Fanuc KAREL source: KT00971.KL

PROGRAM KT00971
%NOLOCKGROUP
VAR
  ENTRY: INTEGER
  PNAME: STRING[80]
  VNAME: STRING[80]
  STATUS: INTEGER
  VALUE: ARRAY[4] OF STRING[20]
BEGIN
  ENTRY = 0
  PNAME = ''
  VNAME = 'VALUE'
  SET_VAR(ENTRY, PNAME, VNAME, VALUE, STATUS)
END KT00971
